Yaskawa INFORM job: 123123.JBI

/JOB
//NAME 123123
//POS
///NPOS 8,8,8,0,0,0
///TOOL 0
///POSTYPE PULSE
///PULSE
C00000=68,-101144,-84203,3631,-80192,-1940
C00001=114331,78034,45532,-5001,-32210,2675
C00002=114374,78891,46569,-5083,-32410,2786
C00003=68,-101145,-84203,3630,-80191,-1940
C00004=130100,113966,38039,100328,-57910,-34898
C00005=125030,110049,33944,101386,-53910,-35608
C00006=126885,100789,21269,102518,-55476,-37189
C00007=131323,99853,36627,90943,-53987,-32131
BC00000=570125
BC00001=756518
BC00002=756937
BC00003=275983
BC00004=275984
BC00005=275984
BC00006=275984
BC00007=275984
EC00000=1491,0
EC00001=7261,0
EC00002=7274,0
EC00003=1491,0
EC00004=1489,0
EC00005=1489,0
EC00006=1489,0
EC00007=1488,0
//INST
///DATE 2023/08/24 12:52
///ATTR SC,RW
///GROUP1 RB1,BS1
///GROUP2 ST2
NOP
MOVJ C00000 BC00000 VJ=90.00  +MOVJ EC00000 VJ=90.00
MOVS C00001 BC00001 V=11.0  +MOVJ EC00001 VJ=0.78
MOVS C00002 BC00002 V=11.0  +MOVJ EC00002 VJ=0.78
MOVJ C00003 BC00003 VJ=90.00  +MOVJ EC00003 VJ=90.00
MOVJ C00004 BC00004 VJ=90.00  +MOVJ EC00004 VJ=90.00
MOVJ C00005 BC00005 VJ=90.00  +MOVJ EC00005 VJ=90.00
MOVL C00006 BC00006 V=1.7  +MOVJ EC00006 VJ=90.00
MOVJ C00007 BC00007 VJ=90.00  +MOVJ EC00007 VJ=90.00
END
